// TIA Portal V19 export
DATA_BLOCK "ACT_SPEED_CS_CP02"   // DB90
// stored: InstanceOfName ACT_SPEED_SCALING, InstanceOfType FB
"ACT_SPEED_SCALING"
   // VAR_INPUT
   //    RAW_MIN : Int;
   //    RAW_MAX : Int;
   //    SCALE_MIN : Real;
   //    SCALE_MAX : Real;
   //    INPUT : Int;
   // END_VAR
   // VAR_OUTPUT
   //    SCALE_OUT : Real;
   // END_VAR
   // VAR
   //    SP : Real;
   // END_VAR
BEGIN
END_DATA_BLOCK
